{attribute 'qualified_only'}
{attribute 'strict'}
{attribute 'to_string'}
TYPE E_Element_State_Short :
(
eNotClean,






eClean,

eProduct




);
END_TYPE

(* stored: Version 1.1.0.1, ProductVersion 3.1.4024.12
   DUT E_Element_State_Short: Id {08b6b406-db46-4dbf-829b-b032e60371d5} *)
